ABB RobotStudio station: MA6212_Projabez.rspag

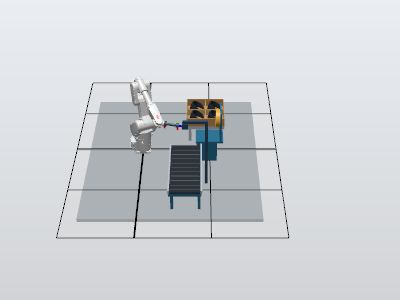
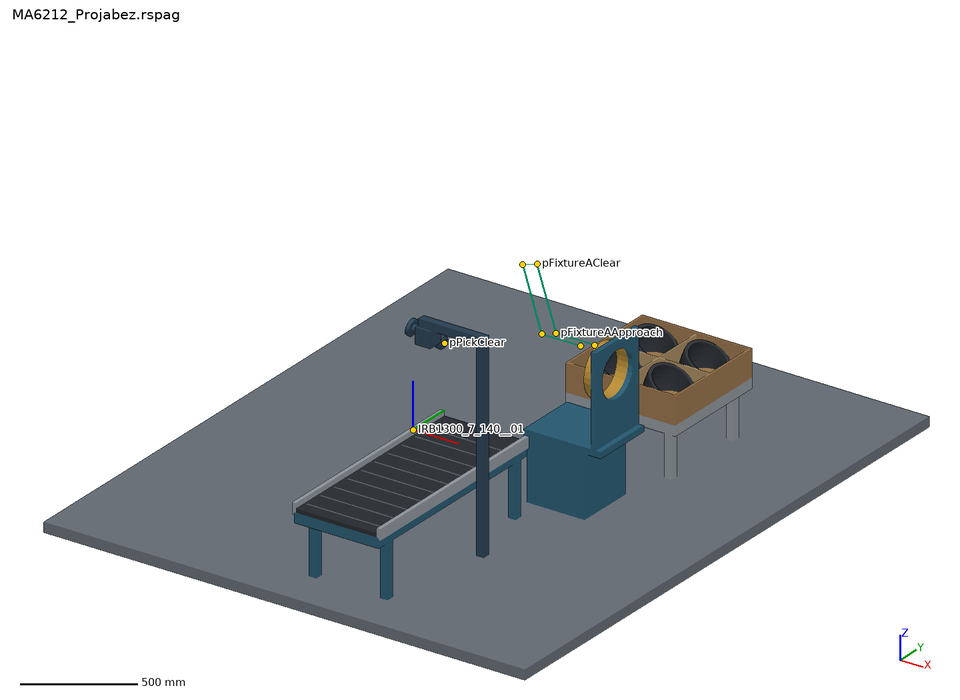
[picture v1: parts stored in the station drawn from their meshes, with robot base, taught points and paths (robot models come from the ABB library and are not in the file)]
--- station ---
Station MA6212_Elbow_Packing (saved by RobotStudio 26.3.11844.1)
Controller MA6212_IRB1300
  mechanical unit ROB_1: IRB1300_7_140__01, 6 joints, base frame (0, 0, 0) mm
Layout (positions relative to the parent item):
  - IRB1300_7_140__01 [mechanism, from %ABB.RobotStudio.Models.IRB1300%\IRB1300_7_140__01.rslib] at (0, 0, 0) mm; joint values [-1.0982, -0.2684, 0.7374, -1.5164, -1.072, 1.13] (rad or m)
  - Cell_Floor [part], size 2500 x 3000 x 50 mm
  - Infeed_Conveyor [part], size 460 x 1100 x 375 mm
  - Gasket_Station [part], size 400 x 320 x 810 mm
  - Packing_Box_2x2 [part], size 570 x 570 x 140 mm
  - Box_Support [part] at (250, 0, 0) mm, size 570 x 570 x 280 mm
  - Vision_Camera [part], size 350 x 80 x 1040 mm
  - Elbow_01 [part] at (1070, 350, 300) mm, size 226.4 x 215 x 150 mm
  - Vacuum_Gripper [part] at (369.79, -550, 813.35) mm, rotated rx 180 ry 80 rz 180 deg, size 80 x 79.6 x 180 mm
  - Elbow_02 [part] at (1070, 620, 299.96) mm, size 226.4 x 215 x 150 mm
  - Elbow_03 [part] at (800, 350, 300.59) mm, size 226.4 x 215 x 150 mm
  - Elbow_04 [part] at (800, 620, 300.19) mm, size 226.4 x 215 x 150 mm
  - Gasket_Reference [part], size 200 x 198.9 x 5 mm
  - Conveyor_Belt_Markers [part] at (0, 7.95, 0) mm, size 390 x 908 x 0.5 mm
  - Fixture_Port [part], size 60 x 258.6 x 260 mm
  - Box_Dividers [part], size 550 x 550 x 110 mm
  - MA6212_PackingSimulation [smart component]
  - Measured_TCP_Trace [part], size 571.5 x 1171.9 x 916.4 mm
Attachment: Vacuum_Gripper is attached to IRB1300_7_140__01 / Link6
Targets, tools, work objects and paths stored in the station and not in the controller backup, written as RAPID:
! task T_ROB1
MODULE Module1
  PROC Preview_Slot1()
    MoveJ pPickClear,v1000,z100,tVac\WObj:=wCell;
    MoveL pPickApproach,v1000,z100,tVac\WObj:=wCell;
    MoveL pPickContact,v1000,z100,tVac\WObj:=wCell;
    MoveL pPickClear,v1000,z100,tVac\WObj:=wCell;
    MoveJ pFixtureAClear,v1000,z100,tVac\WObj:=wCell;
    MoveL pFixtureAApproach,v1000,z100,tVac\WObj:=wCell;
    MoveL pFixtureAContact,v1000,z100,tVac\WObj:=wCell;
    MoveL pFixtureAClear,v1000,z100,tVac\WObj:=wCell;
    MoveJ pFixtureBClear,v1000,z100,tVac\WObj:=wCell;
    MoveL pFixtureBApproach,v1000,z100,tVac\WObj:=wCell;
    MoveL pFixtureBContact,v1000,z100,tVac\WObj:=wCell;
    MoveL pFixtureBClear,v1000,z100,tVac\WObj:=wCell;
    MoveJ pBox1Clear,v1000,z100,tVac\WObj:=wCell;
    MoveL pBox1Approach,v1000,z100,tVac\WObj:=wCell;
    MoveL pBox1Contact,v1000,z100,tVac\WObj:=wCell;
    MoveL pBox1Clear,v1000,z100,tVac\WObj:=wCell;
    MoveJ pPickClear,v1000,z100,tVac\WObj:=wCell;
  ENDPROC
  PROC Preview_Slot2()
    MoveJ pPickClear,v1000,z100,tVac\WObj:=wCell;
    MoveL pPickApproach,v1000,z100,tVac\WObj:=wCell;
    MoveL pPickContact,v1000,z100,tVac\WObj:=wCell;
    MoveL pPickClear,v1000,z100,tVac\WObj:=wCell;
    MoveJ pFixtureAClear,v1000,z100,tVac\WObj:=wCell;
    MoveL pFixtureAApproach,v1000,z100,tVac\WObj:=wCell;
    MoveL pFixtureAContact,v1000,z100,tVac\WObj:=wCell;
    MoveL pFixtureAClear,v1000,z100,tVac\WObj:=wCell;
    MoveJ pFixtureBClear,v1000,z100,tVac\WObj:=wCell;
    MoveL pFixtureBApproach,v1000,z100,tVac\WObj:=wCell;
    MoveL pFixtureBContact,v1000,z100,tVac\WObj:=wCell;
    MoveL pFixtureBClear,v1000,z100,tVac\WObj:=wCell;
    MoveJ pBox2Clear,v1000,z100,tVac\WObj:=wCell;
    MoveL pBox2Approach,v1000,z100,tVac\WObj:=wCell;
    MoveL pBox2Contact,v1000,z100,tVac\WObj:=wCell;
    MoveL pBox2Clear,v1000,z100,tVac\WObj:=wCell;
    MoveJ pPickClear,v1000,z100,tVac\WObj:=wCell;
  ENDPROC
  PROC Preview_Slot3()
    MoveJ pPickClear,v1000,z100,tVac\WObj:=wCell;
    MoveL pPickApproach,v1000,z100,tVac\WObj:=wCell;
    MoveL pPickContact,v1000,z100,tVac\WObj:=wCell;
    MoveL pPickClear,v1000,z100,tVac\WObj:=wCell;
    MoveJ pFixtureAClear,v1000,z100,tVac\WObj:=wCell;
    MoveL pFixtureAApproach,v1000,z100,tVac\WObj:=wCell;
    MoveL pFixtureAContact,v1000,z100,tVac\WObj:=wCell;
    MoveL pFixtureAClear,v1000,z100,tVac\WObj:=wCell;
    MoveJ pFixtureBClear,v1000,z100,tVac\WObj:=wCell;
    MoveL pFixtureBApproach,v1000,z100,tVac\WObj:=wCell;
    MoveL pFixtureBContact,v1000,z100,tVac\WObj:=wCell;
    MoveL pFixtureBClear,v1000,z100,tVac\WObj:=wCell;
    MoveJ pBox3Clear,v1000,z100,tVac\WObj:=wCell;
    MoveL pBox3Approach,v1000,z100,tVac\WObj:=wCell;
    MoveL pBox3Contact,v1000,z100,tVac\WObj:=wCell;
    MoveL pBox3Clear,v1000,z100,tVac\WObj:=wCell;
    MoveJ pPickClear,v1000,z100,tVac\WObj:=wCell;
  ENDPROC
  PROC Preview_Slot4()
    MoveJ pPickClear,v1000,z100,tVac\WObj:=wCell;
    MoveL pPickApproach,v1000,z100,tVac\WObj:=wCell;
    MoveL pPickContact,v1000,z100,tVac\WObj:=wCell;
    MoveL pPickClear,v1000,z100,tVac\WObj:=wCell;
    MoveJ pFixtureAClear,v1000,z100,tVac\WObj:=wCell;
    MoveL pFixtureAApproach,v1000,z100,tVac\WObj:=wCell;
    MoveL pFixtureAContact,v1000,z100,tVac\WObj:=wCell;
    MoveL pFixtureAClear,v1000,z100,tVac\WObj:=wCell;
    MoveJ pFixtureBClear,v1000,z100,tVac\WObj:=wCell;
    MoveL pFixtureBApproach,v1000,z100,tVac\WObj:=wCell;
    MoveL pFixtureBContact,v1000,z100,tVac\WObj:=wCell;
    MoveL pFixtureBClear,v1000,z100,tVac\WObj:=wCell;
    MoveJ pBox4Clear,v1000,z100,tVac\WObj:=wCell;
    MoveL pBox4Approach,v1000,z100,tVac\WObj:=wCell;
    MoveL pBox4Contact,v1000,z100,tVac\WObj:=wCell;
    MoveL pBox4Clear,v1000,z100,tVac\WObj:=wCell;
    MoveJ pPickClear,v1000,z100,tVac\WObj:=wCell;
  ENDPROC
ENDMODULE


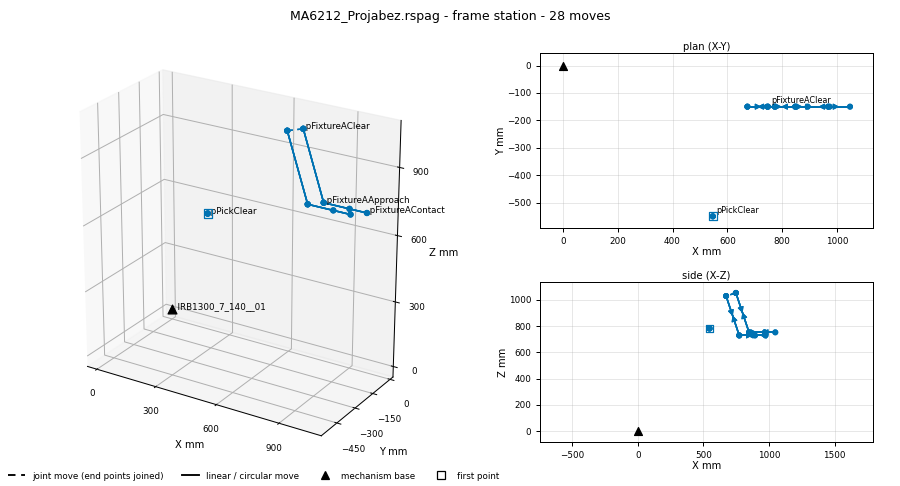
[picture p0: tool path of MA6212_Projabez.rspag in frame station, 28 of 44 moves have a stored position in this frame; points joined in program order, loops and branches not executed]
--- Backups/MA6212_IRB1300/RAPID/TASK1/PROGMOD/MA6212_Packing.modx ---
MODULE MA6212_Packing
    ! Nominal TCP targets: position, orientation, and robot configuration.
    CONST robtarget pPickClear:=[[547.057674,-550,782.094453],[0.642788,-0,0.766044,-0],[-1,-1,0,1],[9E9,9E9,9E9,9E9,9E9,9E9]];
    CONST robtarget pPickApproach:=[[547.057674,-550,562.094453],[0.642788,-0,0.766044,-0],[-1,-1,0,1],[9E9,9E9,9E9,9E9,9E9,9E9]];
    CONST robtarget pPickContact:=[[547.057674,-550,402.094453],[0.642788,-0,0.766044,-0],[-1,-1,0,1],[9E9,9E9,9E9,9E9,9E9,9E9]];
    CONST robtarget pFixtureAClear:=[[747.905547,-150,1052.942326],[0,0.996195,-0,0.087156],[-1,-2,-1,1],[9E9,9E9,9E9,9E9,9E9,9E9]];
    CONST robtarget pFixtureAApproach:=[[847.905547,-150,752.942326],[0,0.996195,-0,0.087156],[-1,-2,-1,1],[9E9,9E9,9E9,9E9,9E9,9E9]];
    CONST robtarget pFixtureAContact:=[[1047.905547,-150,752.942326],[0,0.996195,-0,0.087156],[-1,-2,-1,1],[9E9,9E9,9E9,9E9,9E9,9E9]];
    CONST robtarget pFixtureBClear:=[[673.214521,-150,1029.392336],[0,0.976296,-0,0.21644],[-1,-2,-1,1],[9E9,9E9,9E9,9E9,9E9,9E9]];
    CONST robtarget pFixtureBApproach:=[[773.214521,-150,729.392336],[0,0.976296,-0,0.21644],[-1,-2,-1,1],[9E9,9E9,9E9,9E9,9E9,9E9]];
    CONST robtarget pFixtureBContact:=[[973.214521,-150,729.392336],[0,0.976296,-0,0.21644],[-1,-2,-1,1],[9E9,9E9,9E9,9E9,9E9,9E9]];
    CONST robtarget pBox1Clear:=[[990.607664,350,806.785479],[0.5373,-0,0.843391,-0],[0,1,-2,1],[9E9,9E9,9E9,9E9,9E9,9E9]];
    CONST robtarget pBox1Approach:=[[990.607664,350,586.785479],[0.5373,-0,0.843391,-0],[0,0,-1,1],[9E9,9E9,9E9,9E9,9E9,9E9]];
    CONST robtarget pBox1Contact:=[[990.607664,350,426.785479],[0.5373,-0,0.843391,-0],[0,0,-1,1],[9E9,9E9,9E9,9E9,9E9,9E9]];
    CONST robtarget pBox2Clear:=[[990.607664,620,806.785479],[0.5373,-0,0.843391,-0],[0,1,-2,1],[9E9,9E9,9E9,9E9,9E9,9E9]];
    CONST robtarget pBox2Approach:=[[990.607664,620,586.785479],[0.5373,-0,0.843391,-0],[0,0,-1,1],[9E9,9E9,9E9,9E9,9E9,9E9]];
    CONST robtarget pBox2Contact:=[[990.607664,620,426.785479],[0.5373,-0,0.843391,-0],[0,0,-1,1],[9E9,9E9,9E9,9E9,9E9,9E9]];
    CONST robtarget pBox3Clear:=[[720.607664,350,806.785479],[0.5373,-0,0.843391,-0],[0,1,-2,1],[9E9,9E9,9E9,9E9,9E9,9E9]];
    CONST robtarget pBox3Approach:=[[720.607664,350,586.785479],[0.5373,-0,0.843391,-0],[0,0,-1,1],[9E9,9E9,9E9,9E9,9E9,9E9]];
    CONST robtarget pBox3Contact:=[[720.607664,350,426.785479],[0.5373,-0,0.843391,-0],[0,0,-1,1],[9E9,9E9,9E9,9E9,9E9,9E9]];
    CONST robtarget pBox4Clear:=[[720.607664,620,806.785479],[0.5373,-0,0.843391,-0],[0,1,-1,1],[9E9,9E9,9E9,9E9,9E9,9E9]];
    CONST robtarget pBox4Approach:=[[720.607664,620,586.785479],[0.5373,-0,0.843391,-0],[0,0,-1,1],[9E9,9E9,9E9,9E9,9E9,9E9]];
    CONST robtarget pBox4Contact:=[[720.607664,620,426.785479],[0.5373,-0,0.843391,-0],[0,0,-1,1],[9E9,9E9,9E9,9E9,9E9,9E9]];

    ! Tool, workobject, payload, and shared process variables.
    PERS tooldata tVac:=[TRUE,[[0,0,180],[1,0,0,0]],[1,[0,0,80],[1,0,0,0],0.003,0.003,0.001]];
    PERS wobjdata wCell:=[FALSE,TRUE,"",[[0,0,0],[1,0,0,0]],[[0,0,0],[1,0,0,0]]];
    PERS loaddata loadPipe:=[2.5,[0,0,80],[1,0,0,0],0.02,0.02,0.02];
    PERS num nStage:=50;
    PERS num nPart:=4;
    PERS num nSlot:=4;
    PERS num visionX:=12.7711;
    PERS num visionY:=7.95181;
    PERS num visionYaw:=-4.63855;
    PERS num cycleTimes{4}:=[37.228,38.252,37.088,38.028];
    PERS num totalTime:=150.596;
    PERS bool batchComplete:=TRUE;
    VAR num seed:=317;
    VAR clock cycleClock;
    VAR clock batchClock;
    VAR robtarget pSeen;
    VAR robtarget pBox;

    PROC Stage(num value)
        ! Let the Smart Component observe this process state.
        nStage:=value;
        WaitTime 0.10;
    ENDPROC

    FUNC num RandomUnit()
        seed:=(17*seed+43) MOD 997;
        RETURN seed/996;
    ENDFUNC

    PROC ReadSimulatedVision()
        ! Fixed seed gives repeatable planar offsets and yaw.
        visionX:=30*RandomUnit()-15;
        visionY:=30*RandomUnit()-15;
        visionYaw:=10*RandomUnit()-5;
        pSeen:=pPickContact;
        pSeen.trans.x:=650+visionX-102.942326*Cos(visionYaw);
        pSeen.trans.y:=-550+visionY-102.942326*Sin(visionYaw);
        pSeen.rot:=OrientZYX(visionYaw,100,0);
    ENDPROC

    PROC main()
        ConfJ \On;
        ConfL \Off;
        VelSet 100,800;
        AccSet 60,60;
        batchComplete:=FALSE;
        seed:=317;
        nPart:=0;
        Stage 0;
        GripLoad load0;
        MoveJ pPickClear,v500,fine,tVac\WObj:=wCell;
        ClkReset batchClock;
        ClkStart batchClock;
        FOR partIndex FROM 1 TO 4 DO
            ClkReset cycleClock;
            ClkStart cycleClock;
            ! Clear the previous release stage before updating part identity.
            Stage 5;
            nPart:=partIndex;
            nSlot:=((partIndex-1) MOD 4)+1;
            ReadSimulatedVision;
            ! Index the belt to the pickup position.
            Stage 8;
            WaitTime 3;
            Stage 10;
            ! Pick at contact A and place on the fixture.
            MoveJ Offs(pSeen,0,0,380),v500,z20,tVac\WObj:=wCell;
            MoveL Offs(pSeen,0,0,160),v300,z10,tVac\WObj:=wCell;
            MoveL pSeen,v100,fine,tVac\WObj:=wCell;
            Stage 20;
            GripLoad loadPipe;
            MoveL Offs(pSeen,0,0,380),v200,z10,tVac\WObj:=wCell;
            MoveJ pFixtureAClear,v500,z20,tVac\WObj:=wCell;
            MoveL pFixtureAApproach,v300,z10,tVac\WObj:=wCell;
            MoveL Offs(pFixtureAContact,-80,0,0),v100,fine,tVac\WObj:=wCell;
            ! Insert the inlet into the horizontal wall port.
            Stage 25;
            MoveL pFixtureAContact,v50,fine,tVac\WObj:=wCell;
            Stage 30;
            GripLoad load0;
            MoveL pFixtureAApproach,v100,fine,tVac\WObj:=wCell;
            MoveL pFixtureAClear,v200,fine,tVac\WObj:=wCell;
            ! Gasket machinery is abstracted as a two-second dwell.
            WaitTime 2;
            ! Pick at contact B, then fill the indexed box slot.
            MoveJ pFixtureBClear,v300,fine,tVac\WObj:=wCell;
            MoveL pFixtureBApproach,v200,z10,tVac\WObj:=wCell;
            MoveL pFixtureBContact,v100,fine,tVac\WObj:=wCell;
            Stage 40;
            GripLoad loadPipe;
            ! Withdraw fully before the box transfer.
            MoveL Offs(pFixtureBContact,-80,0,0),v50,fine,tVac\WObj:=wCell;
            Stage 45;
            MoveL pFixtureBApproach,v100,fine,tVac\WObj:=wCell;
            MoveL pFixtureBClear,v200,z10,tVac\WObj:=wCell;
            TEST nSlot
            CASE 1: pBox:=pBox1Contact;
            CASE 2: pBox:=pBox2Contact;
            CASE 3: pBox:=pBox3Contact;
            CASE 4: pBox:=pBox4Contact;
            ENDTEST
            MoveJ Offs(pBox,0,0,380),v500,z20,tVac\WObj:=wCell;
            MoveL Offs(pBox,0,0,160),v200,z10,tVac\WObj:=wCell;
            MoveL pBox,v100,fine,tVac\WObj:=wCell;
            Stage 50;
            GripLoad load0;
            MoveL Offs(pBox,0,0,380),v200,z10,tVac\WObj:=wCell;
            MoveJ pPickClear,v500,fine,tVac\WObj:=wCell;
            ClkStop cycleClock;
            cycleTimes{partIndex}:=ClkRead(cycleClock);
        ENDFOR
        ClkStop batchClock;
        totalTime:=ClkRead(batchClock);
        batchComplete:=TRUE;
        TPWrite "MA6212: 4 parts packed in one divided box.";
    ENDPROC
ENDMODULE

--- Backups/MA6212_IRB1300/HOME/MA6212_Packing.mod ---
MODULE MA6212_Packing
    ! Nominal TCP targets: position, orientation, and robot configuration.
    CONST robtarget pPickClear:=[[547.057674,-550,782.094453],[0.642788,-0,0.766044,-0],[-1,-1,0,1],[9E9,9E9,9E9,9E9,9E9,9E9]];
    CONST robtarget pPickApproach:=[[547.057674,-550,562.094453],[0.642788,-0,0.766044,-0],[-1,-1,0,1],[9E9,9E9,9E9,9E9,9E9,9E9]];
    CONST robtarget pPickContact:=[[547.057674,-550,402.094453],[0.642788,-0,0.766044,-0],[-1,-1,0,1],[9E9,9E9,9E9,9E9,9E9,9E9]];
    CONST robtarget pFixtureAClear:=[[747.905547,-150,1052.942326],[0,0.996195,-0,0.087156],[-1,-2,-1,1],[9E9,9E9,9E9,9E9,9E9,9E9]];
    CONST robtarget pFixtureAApproach:=[[847.905547,-150,752.942326],[0,0.996195,-0,0.087156],[-1,-2,-1,1],[9E9,9E9,9E9,9E9,9E9,9E9]];
    CONST robtarget pFixtureAContact:=[[1047.905547,-150,752.942326],[0,0.996195,-0,0.087156],[-1,-2,-1,1],[9E9,9E9,9E9,9E9,9E9,9E9]];
    CONST robtarget pFixtureBClear:=[[673.214521,-150,1029.392336],[0,0.976296,-0,0.21644],[-1,-2,-1,1],[9E9,9E9,9E9,9E9,9E9,9E9]];
    CONST robtarget pFixtureBApproach:=[[773.214521,-150,729.392336],[0,0.976296,-0,0.21644],[-1,-2,-1,1],[9E9,9E9,9E9,9E9,9E9,9E9]];
    CONST robtarget pFixtureBContact:=[[973.214521,-150,729.392336],[0,0.976296,-0,0.21644],[-1,-2,-1,1],[9E9,9E9,9E9,9E9,9E9,9E9]];
    CONST robtarget pBox1Clear:=[[990.607664,350,806.785479],[0.5373,-0,0.843391,-0],[0,1,-2,1],[9E9,9E9,9E9,9E9,9E9,9E9]];
    CONST robtarget pBox1Approach:=[[990.607664,350,586.785479],[0.5373,-0,0.843391,-0],[0,0,-1,1],[9E9,9E9,9E9,9E9,9E9,9E9]];
    CONST robtarget pBox1Contact:=[[990.607664,350,426.785479],[0.5373,-0,0.843391,-0],[0,0,-1,1],[9E9,9E9,9E9,9E9,9E9,9E9]];
    CONST robtarget pBox2Clear:=[[990.607664,620,806.785479],[0.5373,-0,0.843391,-0],[0,1,-2,1],[9E9,9E9,9E9,9E9,9E9,9E9]];
    CONST robtarget pBox2Approach:=[[990.607664,620,586.785479],[0.5373,-0,0.843391,-0],[0,0,-1,1],[9E9,9E9,9E9,9E9,9E9,9E9]];
    CONST robtarget pBox2Contact:=[[990.607664,620,426.785479],[0.5373,-0,0.843391,-0],[0,0,-1,1],[9E9,9E9,9E9,9E9,9E9,9E9]];
    CONST robtarget pBox3Clear:=[[720.607664,350,806.785479],[0.5373,-0,0.843391,-0],[0,1,-2,1],[9E9,9E9,9E9,9E9,9E9,9E9]];
    CONST robtarget pBox3Approach:=[[720.607664,350,586.785479],[0.5373,-0,0.843391,-0],[0,0,-1,1],[9E9,9E9,9E9,9E9,9E9,9E9]];
    CONST robtarget pBox3Contact:=[[720.607664,350,426.785479],[0.5373,-0,0.843391,-0],[0,0,-1,1],[9E9,9E9,9E9,9E9,9E9,9E9]];
    CONST robtarget pBox4Clear:=[[720.607664,620,806.785479],[0.5373,-0,0.843391,-0],[0,1,-1,1],[9E9,9E9,9E9,9E9,9E9,9E9]];
    CONST robtarget pBox4Approach:=[[720.607664,620,586.785479],[0.5373,-0,0.843391,-0],[0,0,-1,1],[9E9,9E9,9E9,9E9,9E9,9E9]];
    CONST robtarget pBox4Contact:=[[720.607664,620,426.785479],[0.5373,-0,0.843391,-0],[0,0,-1,1],[9E9,9E9,9E9,9E9,9E9,9E9]];

    ! Tool, workobject, payload, and shared process variables.
    PERS tooldata tVac:=[TRUE,[[0,0,180],[1,0,0,0]],[1,[0,0,80],[1,0,0,0],0.003,0.003,0.001]];
    PERS wobjdata wCell:=[FALSE,TRUE,"",[[0,0,0],[1,0,0,0]],[[0,0,0],[1,0,0,0]]];
    PERS loaddata loadPipe:=[2.5,[0,0,80],[1,0,0,0],0.02,0.02,0.02];
    PERS num nStage:=0;
    PERS num nPart:=0;
    PERS num nSlot:=1;
    PERS num visionX:=0;
    PERS num visionY:=0;
    PERS num visionYaw:=0;
    PERS num cycleTimes{4}:=[0,0,0,0];
    PERS num totalTime:=0;
    PERS bool batchComplete:=FALSE;
    VAR num seed:=317;
    VAR clock cycleClock;
    VAR clock batchClock;
    VAR robtarget pSeen;
    VAR robtarget pBox;

    PROC Stage(num value)
        ! Let the Smart Component observe this process state.
        nStage:=value;
        WaitTime 0.10;
    ENDPROC

    FUNC num RandomUnit()
        seed:=(17*seed+43) MOD 997;
        RETURN seed/996;
    ENDFUNC

    PROC ReadSimulatedVision()
        ! Fixed seed gives repeatable planar offsets and yaw.
        visionX:=30*RandomUnit()-15;
        visionY:=30*RandomUnit()-15;
        visionYaw:=10*RandomUnit()-5;
        pSeen:=pPickContact;
        pSeen.trans.x:=650+visionX-102.942326*Cos(visionYaw);
        pSeen.trans.y:=-550+visionY-102.942326*Sin(visionYaw);
        pSeen.rot:=OrientZYX(visionYaw,100,0);
    ENDPROC

    PROC main()
        ConfJ \On;
        ConfL \Off;
        VelSet 100,800;
        AccSet 60,60;
        batchComplete:=FALSE;
        seed:=317;
        nPart:=0;
        Stage 0;
        GripLoad load0;
        MoveJ pPickClear,v500,fine,tVac\WObj:=wCell;
        ClkReset batchClock;
        ClkStart batchClock;
        FOR partIndex FROM 1 TO 4 DO
            ClkReset cycleClock;
            ClkStart cycleClock;
            ! Clear the previous release stage before updating part identity.
            Stage 5;
            nPart:=partIndex;
            nSlot:=((partIndex-1) MOD 4)+1;
            ReadSimulatedVision;
            ! Index the belt to the pickup position.
            Stage 8;
            WaitTime 3;
            Stage 10;
            ! Pick at contact A and place on the fixture.
            MoveJ Offs(pSeen,0,0,380),v500,z20,tVac\WObj:=wCell;
            MoveL Offs(pSeen,0,0,160),v300,z10,tVac\WObj:=wCell;
            MoveL pSeen,v100,fine,tVac\WObj:=wCell;
            Stage 20;
            GripLoad loadPipe;
            MoveL Offs(pSeen,0,0,380),v200,z10,tVac\WObj:=wCell;
            MoveJ pFixtureAClear,v500,z20,tVac\WObj:=wCell;
            MoveL pFixtureAApproach,v300,z10,tVac\WObj:=wCell;
            MoveL Offs(pFixtureAContact,-80,0,0),v100,fine,tVac\WObj:=wCell;
            ! Insert the inlet into the horizontal wall port.
            Stage 25;
            MoveL pFixtureAContact,v50,fine,tVac\WObj:=wCell;
            Stage 30;
            GripLoad load0;
            MoveL pFixtureAApproach,v100,fine,tVac\WObj:=wCell;
            MoveL pFixtureAClear,v200,fine,tVac\WObj:=wCell;
            ! Gasket machinery is abstracted as a two-second dwell.
            WaitTime 2;
            ! Pick at contact B, then fill the indexed box slot.
            MoveJ pFixtureBClear,v300,fine,tVac\WObj:=wCell;
            MoveL pFixtureBApproach,v200,z10,tVac\WObj:=wCell;
            MoveL pFixtureBContact,v100,fine,tVac\WObj:=wCell;
            Stage 40;
            GripLoad loadPipe;
            ! Withdraw fully before the box transfer.
            MoveL Offs(pFixtureBContact,-80,0,0),v50,fine,tVac\WObj:=wCell;
            Stage 45;
            MoveL pFixtureBApproach,v100,fine,tVac\WObj:=wCell;
            MoveL pFixtureBClear,v200,z10,tVac\WObj:=wCell;
            TEST nSlot
            CASE 1: pBox:=pBox1Contact;
            CASE 2: pBox:=pBox2Contact;
            CASE 3: pBox:=pBox3Contact;
            CASE 4: pBox:=pBox4Contact;
            ENDTEST
            MoveJ Offs(pBox,0,0,380),v500,z20,tVac\WObj:=wCell;
            MoveL Offs(pBox,0,0,160),v200,z10,tVac\WObj:=wCell;
            MoveL pBox,v100,fine,tVac\WObj:=wCell;
            Stage 50;
            GripLoad load0;
            MoveL Offs(pBox,0,0,380),v200,z10,tVac\WObj:=wCell;
            MoveJ pPickClear,v500,fine,tVac\WObj:=wCell;
            ClkStop cycleClock;
            cycleTimes{partIndex}:=ClkRead(cycleClock);
        ENDFOR
        ClkStop batchClock;
        totalTime:=ClkRead(batchClock);
        batchComplete:=TRUE;
        TPWrite "MA6212: 4 parts packed in one divided box.";
    ENDPROC
ENDMODULE

--- Backups/MA6212_IRB1300/SYSPAR/EIO.cfg ---
EIO:CFG_1.0:7:0::
#
VIRTUAL_NETWORK:

      -Name "Virtual" -Label "Virtual Device Network"
#
EIO_SIGNAL:

      -Name "IIO_di1" -SignalType "DI" -Device "IntegratedIOInternalDevice"\
      -DeviceMap "0"

      -Name "IIO_di2" -SignalType "DI" -Device "IntegratedIOInternalDevice"\
      -DeviceMap "1"

      -Name "IIO_di3" -SignalType "DI" -Device "IntegratedIOInternalDevice"\
      -DeviceMap "2"

      -Name "IIO_di4" -SignalType "DI" -Device "IntegratedIOInternalDevice"\
      -DeviceMap "3"

      -Name "IIO_di5" -SignalType "DI" -Device "IntegratedIOInternalDevice"\
      -DeviceMap "4"

      -Name "IIO_di6" -SignalType "DI" -Device "IntegratedIOInternalDevice"\
      -DeviceMap "5"

      -Name "IIO_di7" -SignalType "DI" -Device "IntegratedIOInternalDevice"\
      -DeviceMap "6"

      -Name "IIO_di8" -SignalType "DI" -Device "IntegratedIOInternalDevice"\
      -DeviceMap "7"

      -Name "IIO_di9" -SignalType "DI" -Device "IntegratedIOInternalDevice"\
      -DeviceMap "8"

      -Name "IIO_di10" -SignalType "DI" -Device "IntegratedIOInternalDevice"\
      -DeviceMap "9"

      -Name "IIO_di11" -SignalType "DI" -Device "IntegratedIOInternalDevice"\
      -DeviceMap "10"

      -Name "IIO_di12" -SignalType "DI" -Device "IntegratedIOInternalDevice"\
      -DeviceMap "11"

      -Name "IIO_di13" -SignalType "DI" -Device "IntegratedIOInternalDevice"\
      -DeviceMap "12"

      -Name "IIO_di14" -SignalType "DI" -Device "IntegratedIOInternalDevice"\
      -DeviceMap "13"

      -Name "IIO_di15" -SignalType "DI" -Device "IntegratedIOInternalDevice"\
      -DeviceMap "14"

      -Name "IIO_di16" -SignalType "DI" -Device "IntegratedIOInternalDevice"\
      -DeviceMap "15"

      -Name "IIO_do1" -SignalType "DO" -Device "IntegratedIOInternalDevice"\
      -DeviceMap "0"

      -Name "IIO_do2" -SignalType "DO" -Device "IntegratedIOInternalDevice"\
      -DeviceMap "1"

      -Name "IIO_do3" -SignalType "DO" -Device "IntegratedIOInternalDevice"\
      -DeviceMap "2"

      -Name "IIO_do4" -SignalType "DO" -Device "IntegratedIOInternalDevice"\
      -DeviceMap "3"

      -Name "IIO_do5" -SignalType "DO" -Device "IntegratedIOInternalDevice"\
      -DeviceMap "4"

      -Name "IIO_do6" -SignalType "DO" -Device "IntegratedIOInternalDevice"\
      -DeviceMap "5"

      -Name "IIO_do7" -SignalType "DO" -Device "IntegratedIOInternalDevice"\
      -DeviceMap "6"

      -Name "IIO_do8" -SignalType "DO" -Device "IntegratedIOInternalDevice"\
      -DeviceMap "7"

      -Name "IIO_gi" -SignalType "GI" -Device "integratedIOInternalDevice"\
      -DeviceMap "0-15"

      -Name "IIO_go" -SignalType "GO" -Device "integratedIOInternalDevice"\
      -DeviceMap "0-7"

#CTRL_SIGNATURE:qBvZBk7J8xCBBRl1bZzPDkQHFjKT+POykwWBU5wAhTH4dfb2+C0l2PJH4G6KDdh12ckKcgMoJZ+ELTlNrl8irQ==

--- Backups/MA6212_IRB1300/SYSPAR/PROC.cfg ---
PROC:CFG_1.0:7:0::

#CTRL_SIGNATURE:shZx++80xs0VY5e3tzRHzO48SW6tPrFOAyuMrvMI6b8C11Uf9xKfJjnffPSkl4SAObYQMD3NYTsOsuR0RYX5wg==
